FUNCTION_BLOCK FB_CtrlOut_1
(*
Function block used to set output from controller.

Constructor: 		Patryk Panylo
Company:		E. Riexinger GmbH
Date:			03.06.2014
Version:			1.00

Date:			Revision:		Who:				Comment
dd.mm.yyyy		x.xx			Initials			comment

*)
VAR_INPUT
	(* Enummerations *)

	(* Variables *)
	lrInSignal								:LREAL;							(* Input signal *)
	lrSignalOffset							:LREAL := 0.0;						(* Offset signal *)
	lrLimitMin								:LREAL := -1E40;					(* Limit minimum *)
	lrLimitMax							:LREAL := 1E40;					(* Limit maximum *)

	(* References *)

	(* Interfaces *)

	(* Instances *)

END_VAR
VAR_OUTPUT
	(* Enummerations *)

	(* Variables *)
	lrOutSignal							:LREAL;							(* Output signal *)
	bLimitMin							:BOOL;							(* Limit minimum reached *)
	bLimitMax							:BOOL;							(* Limit maximum reached *)

	(* References *)

	(* Interfaces *)

	(* Instances *)
END_VAR
VAR
	(* Enummerations *)

	(* Variables *)

	(* References *)

	(* Interfaces *)

	(* Instances *)
	fbLimiter								:FB_Limiter;						(* Signal output limiter *)

END_VAR


(* Limit the outputs *)
fbLimiter(
	bEnable := TRUE,
	lrInSignal := lrInSignal + lrSignalOffset,
	lrLimitMin := lrLimitMin,
	lrLimitMax := lrLimitMax,
	lrOutSignal => lrOutSignal,
	bLimitMin => bLimitMin,
	bLimitMax => bLimitMax
);

END_FUNCTION_BLOCK

(* stored: Version 1.1.0.1, ProductVersion 3.1.4024.15
   POU FB_CtrlOut_1: Id {dbef6318-9463-4414-97e0-349c4cd76f88}, SpecialFunc None *)
